// TIA Portal V19 export
DATA_BLOCK "SKIDS_DB"   // DB26
// stored: InstanceOfName SKIDS, InstanceOfType FB
"SKIDS"
   // VAR
   //    CHILLED_SKIDS_Instance { S7_SetPoint := 'True'} : "SKIDS_LOGIC";
   //    START_Instance { S7_SetPoint := 'True'} : "START";
   //    START_Instance_COLD_SKIDS { S7_SetPoint := 'True'} : "START";
   //    CS_SKIDS_Instance_1 { S7_SetPoint := 'True'} : "SKIDS_LOGIC";
   //    START_Instance_UCH { S7_SetPoint := 'True'} : "START";
   //    ULTRACHILLED_SKIDS_Instance { S7_SetPoint := 'True'} : "SKIDS_LOGIC";
   //    ULTRACHILLED_SKIDS_Instance_1 { S7_SetPoint := 'True'} : "ULTRACHILLED_SKIDS";
   //    HOT_SKIDS_InstancE { S7_SetPoint := 'True'} : "SKIDS_LOGIC";
   //    HOT_SKIDS_Instance_1 { S7_SetPoint := 'True'} : "HOT_SKIDS";
   //    START_Instance_HOT_SKIDS { S7_SetPoint := 'True'} : "START";
   // END_VAR
BEGIN
END_DATA_BLOCK
